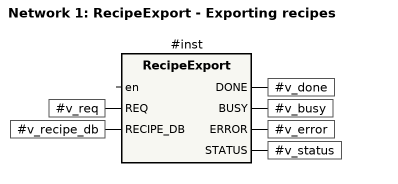
   #inst(REQ := #v_req,   // RecipeExport
         RECIPE_DB := #v_recipe_db,
         DONE => #v_done,
         BUSY => #v_busy,
         ERROR => #v_error,
         STATUS => #v_status);
END_REGION
END_FUNCTION_BLOCK

FUNCTION_BLOCK "FB_Fbd_ex136"   // FB145, FBD
{ S7_Optimized_Access := 'TRUE' }
   VAR_INPUT
      v_req : Bool;
   END_VAR
   VAR_OUTPUT
      v_done : Bool;
      v_busy : Bool;
      v_error : Bool;
      v_status : Word;
   END_VAR
   VAR_IN_OUT
      v_recipe_db : Array[0..99] of Byte;
   END_VAR
   VAR
      inst : RecipeImport;
   END_VAR
BEGIN

REGION Network 1: RecipeImport - Importing recipes
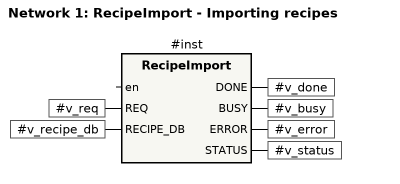
   #inst(REQ := #v_req,   // RecipeImport
         RECIPE_DB := #v_recipe_db,
         DONE => #v_done,
         BUSY => #v_busy,
         ERROR => #v_error,
         STATUS => #v_status);
END_REGION
END_FUNCTION_BLOCK

FUNCTION_BLOCK "FB_Fbd_ex138"   // FB146, FBD
{ S7_Optimized_Access := 'TRUE' }
   VAR_INPUT
      v_req : Bool;
      v_records : UDInt;
      v_format : UInt;
      v_timestamp : UInt;
      v_name : Array[0..99] of Byte;
   END_VAR
   VAR_OUTPUT
      v_done : Bool;
      v_busy : Bool;
      v_error : Bool;
      v_status : Word;
   END_VAR
   VAR_IN_OUT
      v_id : DWord;
      v_header : Array[0..99] of Byte;
      v_data : Array[0..99] of Byte;
   END_VAR
   VAR
      inst : DataLogCreate;
   END_VAR
BEGIN

REGION Network 1: DataLogCreate - Create data log
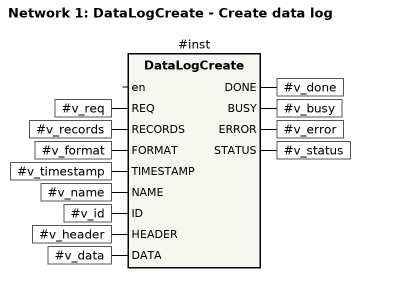
   #inst(REQ := #v_req,   // DataLogCreate
         RECORDS := #v_records,
         FORMAT := #v_format,
         TIMESTAMP := #v_timestamp,
         "NAME" := #v_name,
         ID := #v_id,
         HEADER := #v_header,
         DATA := #v_data,
         DONE => #v_done,
         BUSY => #v_busy,
         ERROR => #v_error,
         STATUS => #v_status);
END_REGION
END_FUNCTION_BLOCK

FUNCTION_BLOCK "FB_Fbd_ex139"   // FB147, FBD
{ S7_Optimized_Access := 'TRUE' }
   VAR_INPUT
      v_req : Bool;
      v_mode : UInt;
      v_name : Array[0..99] of Byte;
   END_VAR
   VAR_OUTPUT
      v_done : Bool;
      v_busy : Bool;
      v_error : Bool;
      v_status : Word;
   END_VAR
   VAR_IN_OUT
      v_id : DWord;
      v_data : Variant;
   END_VAR
   VAR
      inst : DataLogOpen;
   END_VAR
BEGIN

REGION Network 1: DataLogOpen - Open data log
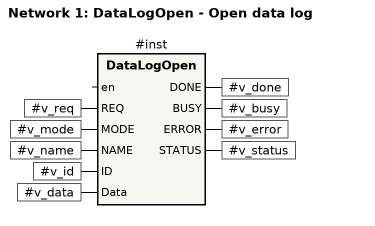
   #inst(REQ := #v_req,   // DataLogOpen
         MODE := #v_mode,
         "NAME" := #v_name,
         ID := #v_id,
         Data := #v_data,
         DONE => #v_done,
         BUSY => #v_busy,
         ERROR => #v_error,
         STATUS => #v_status);
END_REGION
END_FUNCTION_BLOCK

FUNCTION_BLOCK "FB_Fbd_ex140"   // FB148, FBD
{ S7_Optimized_Access := 'TRUE' }
   VAR_INPUT
      v_req : Bool;
      v_mode : UInt;
      v_name : Array[0..99] of Byte;
   END_VAR
   VAR_OUTPUT
      v_done : Bool;
      v_busy : Bool;
      v_error : Bool;
      v_status : Word;
   END_VAR
   VAR_IN_OUT
      v_id : DWord;
      v_data : Array[0..99] of Byte;
   END_VAR
   VAR
      inst : DataLogOpen;
   END_VAR
BEGIN

REGION Network 1: DataLogOpen - Open data log
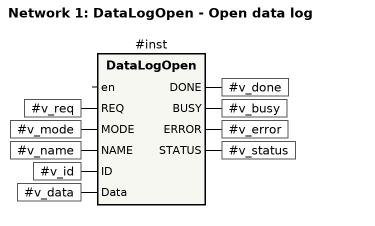
   #inst(REQ := #v_req,   // DataLogOpen
         MODE := #v_mode,
         "NAME" := #v_name,
         ID := #v_id,
         Data := #v_data,
         DONE => #v_done,
         BUSY => #v_busy,
         ERROR => #v_error,
         STATUS => #v_status);
END_REGION
END_FUNCTION_BLOCK

FUNCTION_BLOCK "FB_Fbd_ex141"   // FB149, FBD
{ S7_Optimized_Access := 'TRUE' }
   VAR_INPUT
      v_req : Bool;
   END_VAR
   VAR_OUTPUT
      v_done : Bool;
      v_busy : Bool;
      v_error : Bool;
      v_status : Word;
   END_VAR
   VAR_IN_OUT
      v_id : DWord;
   END_VAR
   VAR
      inst : DataLogClear;
   END_VAR
BEGIN

REGION Network 1: DataLogClear - Empty data log
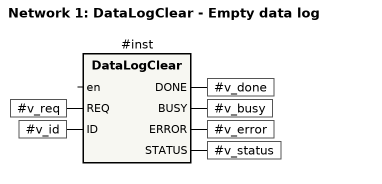
   #inst(REQ := #v_req, ID := #v_id, DONE => #v_done, BUSY => #v_busy, ERROR => #v_error, STATUS => #v_status);   // DataLogClear
END_REGION
END_FUNCTION_BLOCK

FUNCTION_BLOCK "FB_Fbd_ex142"   // FB150, FBD
{ S7_Optimized_Access := 'TRUE' }
   VAR_INPUT
      v_req : Bool;
   END_VAR
   VAR_OUTPUT
      v_done : Bool;
      v_busy : Bool;
      v_error : Bool;
      v_status : Word;
   END_VAR
   VAR_IN_OUT
      v_id : DWord;
   END_VAR
   VAR
      inst : DataLogWrite;
   END_VAR
BEGIN

REGION Network 1: DataLogWrite - Write data log
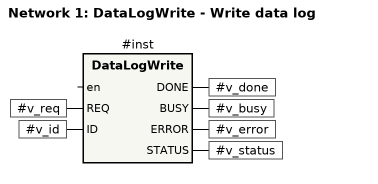
   #inst(REQ := #v_req, ID := #v_id, DONE => #v_done, BUSY => #v_busy, ERROR => #v_error, STATUS => #v_status);   // DataLogWrite
END_REGION
END_FUNCTION_BLOCK

FUNCTION_BLOCK "FB_Fbd_ex143"   // FB151, FBD
{ S7_Optimized_Access := 'TRUE' }
   VAR_INPUT
      v_req : Bool;
   END_VAR
   VAR_OUTPUT
      v_done : Bool;
      v_busy : Bool;
      v_error : Bool;
      v_status : Word;
   END_VAR
   VAR_IN_OUT
      v_id : DWord;
   END_VAR
   VAR
      inst : DataLogClose;
   END_VAR
BEGIN

REGION Network 1: DataLogClose - Close data log
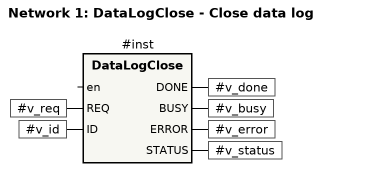
   #inst(REQ := #v_req, ID := #v_id, DONE => #v_done, BUSY => #v_busy, ERROR => #v_error, STATUS => #v_status);   // DataLogClose
END_REGION
END_FUNCTION_BLOCK

FUNCTION_BLOCK "FB_Fbd_ex144"   // FB152, FBD
{ S7_Optimized_Access := 'TRUE' }
   VAR_INPUT
      v_req : Bool;
      v_name : Array[0..99] of Byte;
      v_delfile : Bool;
   END_VAR
   VAR_OUTPUT
      v_done : Bool;
      v_busy : Bool;
      v_error : Bool;
      v_status : Word;
   END_VAR
   VAR_IN_OUT
      v_id : DWord;
   END_VAR
   VAR
      inst : DataLogDelete;
   END_VAR
BEGIN

REGION Network 1: DataLogDelete - Delete data log
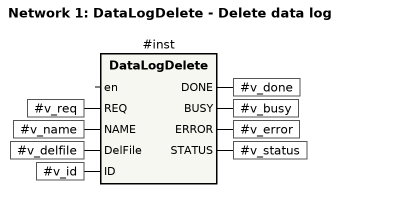
   #inst(REQ := #v_req,   // DataLogDelete
         "NAME" := #v_name,
         DelFile := #v_delfile,
         ID := #v_id,
         DONE => #v_done,
         BUSY => #v_busy,
         ERROR => #v_error,
         STATUS => #v_status);
END_REGION
END_FUNCTION_BLOCK

FUNCTION_BLOCK "FB_Fbd_ex145"   // FB153, FBD
{ S7_Optimized_Access := 'TRUE' }
   VAR_INPUT
      v_req : Bool;
      v_records : UDInt;
      v_name : Array[0..99] of Byte;
   END_VAR
   VAR_OUTPUT
      v_done : Bool;
      v_busy : Bool;
      v_error : Bool;
      v_status : Word;
   END_VAR
   VAR_IN_OUT
      v_id : DWord;
      v_data : Variant;
   END_VAR
   VAR
      inst : DataLogNewFile;
   END_VAR
BEGIN

REGION Network 1: DataLogNewFile - Data log in new file
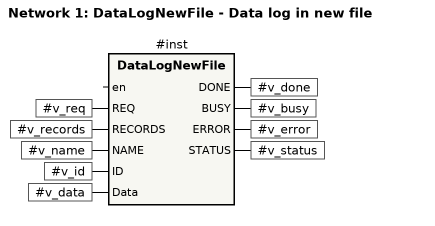
   #inst(REQ := #v_req,   // DataLogNewFile
         RECORDS := #v_records,
         "NAME" := #v_name,
         ID := #v_id,
         Data := #v_data,
         DONE => #v_done,
         BUSY => #v_busy,
         ERROR => #v_error,
         STATUS => #v_status);
END_REGION
END_FUNCTION_BLOCK

FUNCTION_BLOCK "FB_Fbd_ex146"   // FB154, FBD
{ S7_Optimized_Access := 'TRUE' }
   VAR_INPUT
      v_req : Bool;
      v_records : UDInt;
      v_name : Array[0..99] of Byte;
   END_VAR
   VAR_OUTPUT
      v_done : Bool;
      v_busy : Bool;
      v_error : Bool;
      v_status : Word;
   END_VAR
   VAR_IN_OUT
      v_id : DWord;
      v_data : Array[0..99] of Byte;
   END_VAR
   VAR
      inst : DataLogNewFile;
   END_VAR
BEGIN

REGION Network 1: DataLogNewFile - Data log in new file
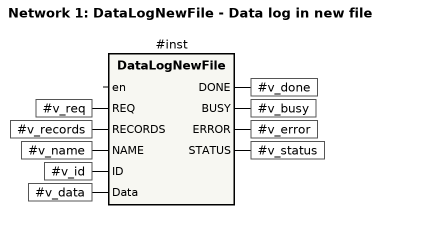
   #inst(REQ := #v_req,   // DataLogNewFile
         RECORDS := #v_records,
         "NAME" := #v_name,
         ID := #v_id,
         Data := #v_data,
         DONE => #v_done,
         BUSY => #v_busy,
         ERROR => #v_error,
         STATUS => #v_status);
END_REGION
END_FUNCTION_BLOCK

FUNCTION_BLOCK "FB_Fbd_ex147"   // FB155, FBD
{ S7_Optimized_Access := 'TRUE' }
   VAR_INPUT
      v_req : Bool;
      v_low_limit : UInt;
      v_up_limit : UInt;
      v_count : UDInt;
      v_attrib : Byte;
      v_srcblk : Variant;
   END_VAR
   VAR_OUTPUT
      v_ret_val : Int;
      v_busy : Bool;
      v_db_num : UInt;
   END_VAR
BEGIN

REGION Network 1: CREATE_DB - Create data block
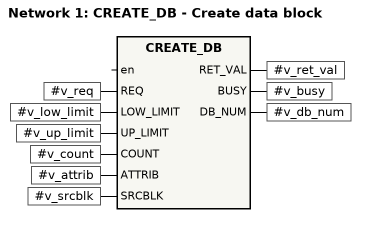
   #v_ret_val := CREATE_DB(REQ := #v_req,
                           LOW_LIMIT := #v_low_limit,
                           UP_LIMIT := #v_up_limit,
                           COUNT := #v_count,
                           ATTRIB := #v_attrib,
                           SRCBLK := #v_srcblk,
                           BUSY => #v_busy,
                           DB_NUM => #v_db_num);
END_REGION
END_FUNCTION_BLOCK

FUNCTION_BLOCK "FB_Fbd_ex148"   // FB156, FBD
{ S7_Optimized_Access := 'TRUE' }
   VAR_INPUT
      v_req : Bool;
   END_VAR
   VAR_OUTPUT
      v_ret_val : Int;
      v_busy : Bool;
   END_VAR
   VAR_IN_OUT
      v_srcblk : Variant;
      v_dstblk : Variant;
   END_VAR
BEGIN

REGION Network 1: READ_DBL - Read from data block in the load memory
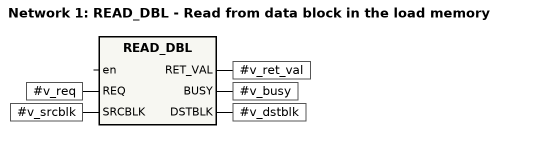
   #v_ret_val := READ_DBL(REQ := #v_req, SRCBLK := #v_srcblk, BUSY => #v_busy, DSTBLK => #v_dstblk);
END_REGION
END_FUNCTION_BLOCK

FUNCTION_BLOCK "FB_Fbd_ex149"   // FB157, FBD
{ S7_Optimized_Access := 'TRUE' }
   VAR_INPUT
      v_req : Bool;
   END_VAR
   VAR_OUTPUT
      v_ret_val : Int;
      v_busy : Bool;
   END_VAR
   VAR_IN_OUT
      v_srcblk : Variant;
      v_dstblk : Variant;
   END_VAR
BEGIN

REGION Network 1: WRIT_DBL - Write to data block in the load memory
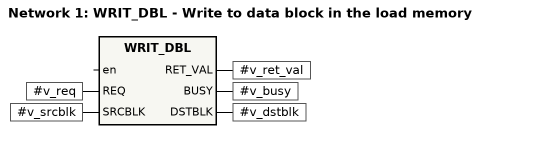
   #v_ret_val := WRIT_DBL(REQ := #v_req, SRCBLK := #v_srcblk, BUSY => #v_busy, DSTBLK => #v_dstblk);
END_REGION
END_FUNCTION_BLOCK

FUNCTION_BLOCK "FB_Fbd_ex150"   // FB158, FBD
{ S7_Optimized_Access := 'TRUE' }
   VAR_INPUT
      v_req : Bool;
      v_db_number : DB_ANY;
   END_VAR
   VAR_OUTPUT
      v_ret_val : Int;
      v_db_length : UDInt;
      v_attrib : Byte;
   END_VAR
BEGIN

REGION Network 1: ATTR_DB - Read data block attribute
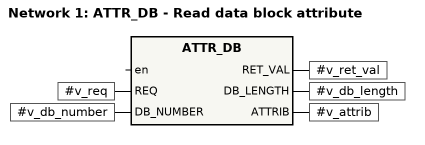
   #v_ret_val := ATTR_DB(REQ := #v_req,
                         DB_NUMBER := #v_db_number,
                         DB_LENGTH => #v_db_length,
                         ATTRIB => #v_attrib);
END_REGION
END_FUNCTION_BLOCK

FUNCTION_BLOCK "FB_Fbd_ex151"   // FB159, FBD
{ S7_Optimized_Access := 'TRUE' }
   VAR_INPUT
      v_req : Bool;
      v_db_number : UInt;
   END_VAR
   VAR_OUTPUT
      v_ret_val : Int;
      v_busy : Bool;
   END_VAR
BEGIN

REGION Network 1: DELETE_DB - Delete data block
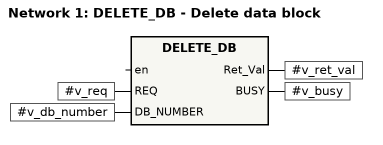
   #v_ret_val := DELETE_DB(REQ := #v_req, DB_NUMBER := #v_db_number, BUSY => #v_busy);
END_REGION
END_FUNCTION_BLOCK

FUNCTION_BLOCK "FB_Fbd_ex152"   // FB160, FBD
{ S7_Optimized_Access := 'TRUE' }
   VAR_INPUT
      v_geoaddr : GEOADDR;
   END_VAR
   VAR_OUTPUT
      v_ret_val : Int;
      v_laddr : UInt;
   END_VAR
BEGIN

REGION Network 1: GEO2LOG - Determine hardware identifier from slot
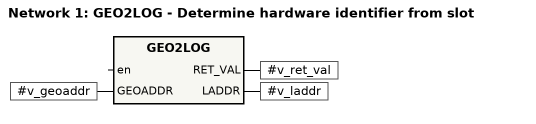
   #v_ret_val := GEO2LOG(GEOADDR := #v_geoaddr, LADDR => #v_laddr);
END_REGION
END_FUNCTION_BLOCK

FUNCTION_BLOCK "FB_Fbd_ex153"   // FB161, FBD
{ S7_Optimized_Access := 'TRUE' }
   VAR_INPUT
      v_laddr : Hw_Any;
   END_VAR
   VAR_OUTPUT
      v_ret_val : Int;
   END_VAR
   VAR_IN_OUT
      v_geoaddr : GEOADDR;
   END_VAR
BEGIN

REGION Network 1: LOG2GEO - Determine slot from hardware identifier
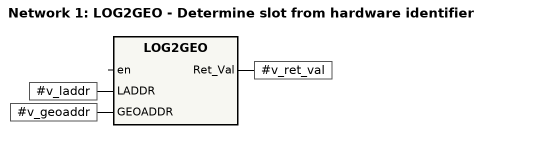
   #v_ret_val := LOG2GEO(LADDR := #v_laddr, GEOADDR := #v_geoaddr);
END_REGION
END_FUNCTION_BLOCK

FUNCTION_BLOCK "FB_Fbd_ex154"   // FB162, FBD
{ S7_Optimized_Access := 'TRUE' }
   VAR_INPUT
      v_ioid : Byte;
      v_addr : Word;
   END_VAR
   VAR_OUTPUT
      v_ret_val : Int;
      v_hwid : Hw_Io;
   END_VAR
BEGIN

REGION Network 1: LOG2MOD - Determine the hardware identifier from addressing of STEP 7 V5.5 SPx
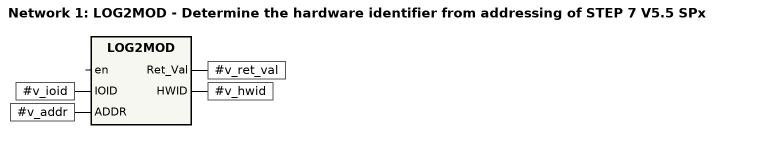
   #v_ret_val := LOG2MOD(IOID := #v_ioid, ADDR := #v_addr, HWID => #v_hwid);
END_REGION
END_FUNCTION_BLOCK

FUNCTION_BLOCK "FB_Fbd_ex155"   // FB163, FBD
{ S7_Optimized_Access := 'TRUE' }
   VAR_INPUT
      v_addr : Variant;
   END_VAR
   VAR_OUTPUT
      v_ret_val : Int;
      v_laddr : Hw_Io;
   END_VAR
BEGIN

REGION Network 1: IO2MOD - Determine hardware identifier from an IO address
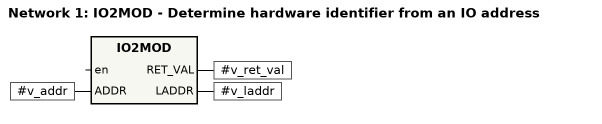
   #v_ret_val := IO2MOD(ADDR := #v_addr, LADDR => #v_laddr);
END_REGION
END_FUNCTION_BLOCK

FUNCTION_BLOCK "FB_Fbd_ex156"   // FB164, FBD
{ S7_Optimized_Access := 'TRUE' }
   VAR_INPUT
      v_laddr : Hw_Io;
   END_VAR
   VAR_OUTPUT
      v_ret_val : Int;
      v_piaddr : UDInt;
      v_picount : UInt;
      v_pqaddr : UDInt;
      v_pqcount : UInt;
   END_VAR
BEGIN

REGION Network 1: RD_ADDR - Determine IO addresses from the hardware identifier
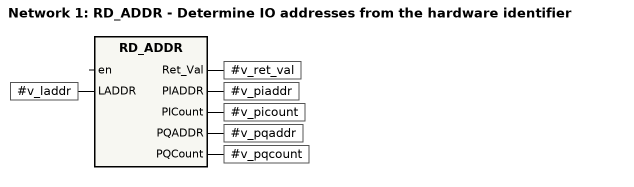
   #v_ret_val := RD_ADDR(LADDR := #v_laddr,
                         PIADDR => #v_piaddr,
                         PICount => #v_picount,
                         PQADDR => #v_pqaddr,
                         PQCount => #v_pqcount);
END_REGION
END_FUNCTION_BLOCK

FUNCTION_BLOCK "FB_Fbd_ex157"   // FB165, FBD
{ S7_Optimized_Access := 'TRUE' }
   VAR_INPUT
      v_master : Int;
      v_station : Int;
      v_slot : Int;
      v_subslot : Int;
   END_VAR
   VAR_OUTPUT
      v_ret_val : Int;
      v_laddr : Hw_Io;
   END_VAR
BEGIN

REGION Network 1: GEO_LOG - Determine hardware identifier from slot
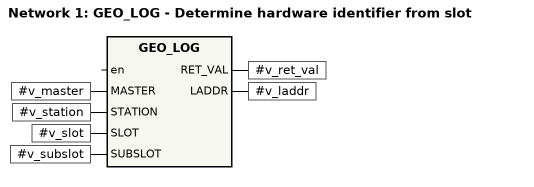
   #v_ret_val := GEO_LOG(MASTER := #v_master,
                         STATION := #v_station,
                         SLOT := #v_slot,
                         SUBSLOT := #v_subslot,
                         LADDR => #v_laddr);
END_REGION
END_FUNCTION_BLOCK

FUNCTION_BLOCK "FB_Fbd_ex158"   // FB166, FBD
{ S7_Optimized_Access := 'TRUE' }
   VAR_INPUT
      v_laddr : Hw_Io;
   END_VAR
   VAR_OUTPUT
      v_ret_val : Int;
      v_area : Int;
      v_master : Int;
      v_station : Int;
      v_slot : Int;
      v_subslot : Int;
      v_offset : Int;
   END_VAR
BEGIN

REGION Network 1: LOG_GEO - Determine slot from hardware identifier
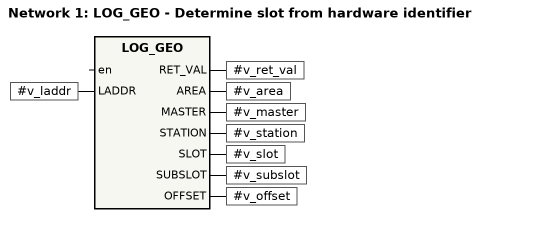
   #v_ret_val := LOG_GEO(LADDR := #v_laddr,
                         AREA => #v_area,
                         MASTER => #v_master,
                         STATION => #v_station,
                         SLOT => #v_slot,
                         SUBSLOT => #v_subslot,
                         OFFSET => #v_offset);
END_REGION
END_FUNCTION_BLOCK

FUNCTION_BLOCK "FB_Fbd_ex160"   // FB167, FBD
{ S7_Optimized_Access := 'TRUE' }
   VAR_INPUT
      v_subnetid : Byte;
      v_rack : Word;
      v_slot : Word;
      v_subslot : Byte;
      v_subaddr : Word;
   END_VAR
   VAR_OUTPUT
      v_ret_val : Int;
      v_ioid : Byte;
      v_laddr : Hw_Module;
   END_VAR
BEGIN

REGION Network 1: GADR_LGC - Determine hardware identifier from slot and offset in the user data address area
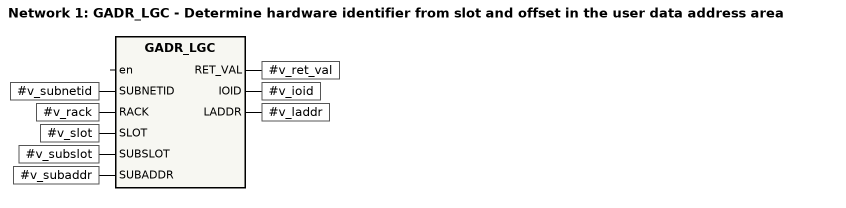
   #v_ret_val := GADR_LGC(SUBNETID := #v_subnetid,
                          RACK := #v_rack,
                          SLOT := #v_slot,
                          SUBSLOT := #v_subslot,
                          SUBADDR := #v_subaddr,
                          IOID => #v_ioid,
                          LADDR => #v_laddr);
END_REGION
END_FUNCTION_BLOCK

FUNCTION_BLOCK "FB_Fbd_ex161"   // FB168, FBD
{ S7_Optimized_Access := 'TRUE' }
   VAR_INPUT
      v_ioid : Byte;
      v_laddr : Hw_Module;
   END_VAR
   VAR_OUTPUT
      v_ret_val : Int;
      v_area : Byte;
      v_rack : Word;
      v_slot : Word;
      v_subaddr : Word;
   END_VAR
BEGIN

REGION Network 1: LGC_GADR - Determine slot from hardware identifier
